# EPICS IOC start-up script: examples/test/PSI/ep2008.iocsh
#- #############################################################################
#- mXsXXX naming
require ecmccfg, "NAMING=mXsXXX"

#- add slaves
${SCRIPTEXEC} ${ecmccfg_DIR}addSlave.cmd, "HW_DESC=EP2008, SLAVE_ID=4"
